(* IEC 61131-3 sources: llm-plc-st-eval/data/processed_definitivo/gpt-4o-2024-08-06/B7/zero_shot, 3 files *)

(* ---- ejec_2.st ---- *)
FUNCTION_BLOCK SelBomba
VAR_INPUT
    modoAuto : BOOL;    // Indica si el modo automático está activo
    btnManual : BOOL;   // Estado del botón manual
    nivelBajo : BOOL;   // Indica si el nivel bajo está activo
END_VAR

VAR_OUTPUT
    bomba : BOOL;       // Estado de la bomba
END_VAR

// Lógica de control de la bomba
// Si modo automático está activo, la bomba se enciende si nivelBajo está activo
// Si modo automático no está activo, la bomba sigue el estado del botón manual
bomba := (modoAuto AND nivelBajo) OR (NOT modoAuto AND btnManual);

END_FUNCTION_BLOCK

(* ---- ejec_3.st ---- *)
FUNCTION_BLOCK SelBomba
VAR_INPUT
    modoAuto : BOOL;    // Indica si el modo automático está activo
    btnManual : BOOL;   // Estado del botón manual
    nivelBajo : BOOL;   // Indica si el nivel bajo está activo
END_VAR
VAR_OUTPUT
    bomba : BOOL;       // Estado de la bomba
END_VAR

// Lógica de control de la bomba
bomba := (modoAuto AND nivelBajo) OR (NOT modoAuto AND btnManual);

END_FUNCTION_BLOCK

(* ---- ejec_1.st ---- *)
PROGRAM SelBomba
VAR
    modoAuto : BOOL;    // Entrada: selecciona el modo automático
    btnManual : BOOL;   // Entrada: botón manual para encender la bomba
    nivelBajo : BOOL;   // Entrada: indica si el nivel es bajo
    bomba : BOOL;       // Salida: estado de la bomba
END_VAR

// Lógica de selección de la fuente de mando de la bomba
IF modoAuto THEN
    // Modo automático: la bomba se enciende si nivelBajo está activo
    bomba := nivelBajo;
ELSE
    // Modo manual: la bomba sigue el estado del botón manual
    bomba := btnManual;
END_IF;
